SUBAPPLICATION logiBUS_AI_Calibrate_3P_OPC (* logiBUS_AI 3-Punkt-Kalibrierung, INI-persistiert, C_MIN/C_MID/C_MAX per Methode, alles per OPC-UA (ohne VT) *)
  (* Standard: 61499-2; Description: Copyright (c) 2026 Meisterschulen am Ostbahnhof This program and the accompanying materials are made available under the terms of the Eclipse Public License 2.0 which is available at https://www.eclipse.org/legal/epl-2.0/ SPDX-License-Identifier: EPL-2.0 *)
  (* Version 1.2, 2026-11-25, Franz Höpfinger, Meisterschulen am Ostbahnhof, SERVER_0 -> MyLib::net::SERVER_0_QO (IND nur bei QO=TRUE, RSP intern). Ein gescheitertes RSP meldet IND mit QO=FALSE, direkt IND->RSP ergab eine Endlosschleife. *)
  (* Version 1.1, 2026-11-04, Franz Höpfinger, Meisterschulen am Ostbahnhof, Neuer optionaler Ausgangs-Plug CAL_OUT (kalibrierter Wert = CALIBRATE.Y, AR) per AR_SPLIT_2 SplitCal zwischen CALIBRATE.Y und PublishCal - wie CAL_OUT in logiBUS_AI_Calibrate_3P_Remote_IDA_OPC. Damit kann z.B. ein Servo direkt am kalibrierten Wert haengen statt den eigenen OPC-UA-Knoten lokal zu abonnieren. Unverdrahtet lassen, wenn nicht gebraucht. *)
  (* Version 1.0, 2026-10-28, Franz Höpfinger, Meisterschulen am Ostbahnhof, Kopie von MyLib::sys::logiBUS_AI_Calibrate_3P_IDA_OPC (INIT-Kette Stand bf9ac7c9) ohne VT, fuer Stationen ohne VT (keine isobus_UT-Libs). InputRaw -> MyLib::sys::logiBUS_AI_Raw_AR_OPC, *_REF_LIT -> MyLib::sys::OPC_TO_AR2, Trigger* -> SERVER_0 (IND->RSP), Publish* -> MyLib::sys::AR_TO_Publish_OPC. VT-Objekt-Parameter entfallen, Kalibrierlogik und INI-Keys unveraendert. *)
  PACKAGE MyLib::sys;
  IMPORT logiBUS::io::AI::logiBUS_AI;
  IMPORT logiBUS::io::AI::logiBUS_AI_S;
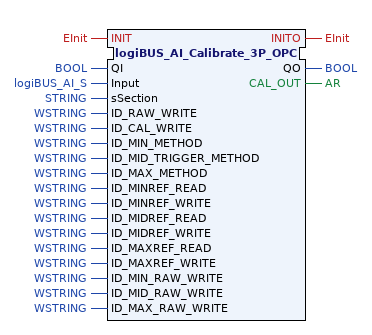
  EVENT_INPUT
    INIT : EInit; (* Initialization Request *)
  END_EVENT
  EVENT_OUTPUT
    INITO : EInit; (* Initialization Confirm *)
  END_EVENT
  VAR_INPUT
    QI : BOOL := TRUE; (* Quality Input - TRUE to enable service *)
    Input : logiBUS::io::AI::logiBUS_AI_S := logiBUS_AI::Invalid; (* Identify the Input AnalogInput_I1..I8 *)
    sSection : STRING; (* INI-Sektionsname fuer X_MIN/X_MID/X_MAX/MIN_REF/MID_REF/MAX_REF-Persistenz - pro Kanal eindeutig, sonst kollidieren die Kanaele in settings.ini *)
    ID_RAW_WRITE : WSTRING; (* Rohwert-Ruckmelde-Adresse (DWORD 0-4095, ACTION=PUBLISH) *)
    ID_CAL_WRITE : WSTRING; (* Kalibrierter-Wert-Ruckmelde-Adresse (REAL, ACTION=PUBLISH) *)
    ID_MIN_METHOD : WSTRING; (* Methodenadresse (ACTION=CREATE_METHOD) fuer den argumentlosen C_MIN-Trigger - gleichberechtigt zur lokalen VT-Taste aufrufbar, sowohl vom OPC-UA-Dashboard als auch per CLIENT_0 von einer anderen Station (siehe OPC_UA_VERNETZUNG.md Punkt 14 - kein Toggle/Subscribe-Umweg mehr) *)
    ID_MID_TRIGGER_METHOD : WSTRING; (* Methodenadresse (ACTION=CREATE_METHOD) fuer den argumentlosen C_MID-Trigger - siehe ID_MIN_METHOD *)
    ID_MAX_METHOD : WSTRING; (* Methodenadresse (ACTION=CREATE_METHOD) fuer den argumentlosen C_MAX-Trigger - siehe ID_MIN_METHOD *)
    ID_MINREF_READ : WSTRING; (* Remote-Subscribe-Adresse MIN_REF-Referenzwert (REAL, ACTION=SUBSCRIBE) *)
    ID_MINREF_WRITE : WSTRING; (* Remote-Echo-Adresse MIN_REF-Referenzwert (REAL, ACTION=PUBLISH) *)
    ID_MIDREF_READ : WSTRING; (* Remote-Subscribe-Adresse MID_REF-Referenzwert (REAL, ACTION=SUBSCRIBE) *)
    ID_MIDREF_WRITE : WSTRING; (* Remote-Echo-Adresse MID_REF-Referenzwert (REAL, ACTION=PUBLISH) *)
    ID_MAXREF_READ : WSTRING; (* Remote-Subscribe-Adresse MAX_REF-Referenzwert (REAL, ACTION=SUBSCRIBE) *)
    ID_MAXREF_WRITE : WSTRING; (* Remote-Echo-Adresse MAX_REF-Referenzwert (REAL, ACTION=PUBLISH) *)
    ID_MIN_RAW_WRITE : WSTRING; (* Rohwert-am-MIN-Kalibrierpunkt-Publish-Adresse (REAL, ACTION=PUBLISH) *)
    ID_MID_RAW_WRITE : WSTRING; (* Rohwert-am-MID-Kalibrierpunkt-Publish-Adresse (REAL, ACTION=PUBLISH) *)
    ID_MAX_RAW_WRITE : WSTRING; (* Rohwert-am-MAX-Kalibrierpunkt-Publish-Adresse (REAL, ACTION=PUBLISH) *)
  END_VAR
  VAR_OUTPUT
    QO : BOOL; (* Quality Output - TRUE if service executed successfully *)
  END_VAR
  PLUGS
    CAL_OUT : adapter::types::unidirectional::AR; (* Optional: kalibrierter Wert (= CALIBRATE.Y) fuer externe Consumer, statt eigenem lokalen OPC-UA-Self-Subscribe auf ID_CAL_WRITE. Unverdrahtet lassen, wenn nicht gebraucht. *)
  END_PLUGS
  FBS
    CALIBRATE : adapter::Engineering::measurements::AR_CALIBRATE_3P_REF(xClipping := FALSE);
    INI_X_MIN : eclipse4diac::storage::INI_AR2(SETM := TRUE, KEY := 'X_MIN', DEFAULT_VALUE := REAL#0.0);
    INI_X_MID : eclipse4diac::storage::INI_AR2(SETM := TRUE, KEY := 'X_MID', DEFAULT_VALUE := REAL#0.0);
    INI_X_MAX : eclipse4diac::storage::INI_AR2(SETM := TRUE, KEY := 'X_MAX', DEFAULT_VALUE := REAL#0.0);
    INI_MIN_REF : eclipse4diac::storage::INI_AR2(SETM := TRUE, KEY := 'MIN_REF', DEFAULT_VALUE := REAL#-100.0);
    INI_MID_REF : eclipse4diac::storage::INI_AR2(SETM := TRUE, KEY := 'MID_REF', DEFAULT_VALUE := REAL#0.0);
    INI_MAX_REF : eclipse4diac::storage::INI_AR2(SETM := TRUE, KEY := 'MAX_REF', DEFAULT_VALUE := REAL#100.0);
    TapMinRaw : adapter::events::bidirectional::AR2_SPLIT_FWD_REV;
    TapMidRaw : adapter::events::bidirectional::AR2_SPLIT_FWD_REV;
    TapMaxRaw : adapter::events::bidirectional::AR2_SPLIT_FWD_REV;
    AND_QO : iec61131::booleanOperators::AND_BOOL_18;
    SplitCal : adapter::events::unidirectional::AR_SPLIT_2;
  END_FBS
  SUBAPPS
    InputRaw : MyLib::sys::logiBUS_AI_Raw_AR_OPC;
    MIN_REF_LIT : MyLib::sys::OPC_TO_AR2;
    MID_REF_LIT : MyLib::sys::OPC_TO_AR2;
    MAX_REF_LIT : MyLib::sys::OPC_TO_AR2;
    TriggerMIN : MyLib::net::SERVER_0_QO; (* RSP direkt auf IND (sonst 4s Server-Lock) *)
    TriggerMID : MyLib::net::SERVER_0_QO; (* RSP direkt auf IND (sonst 4s Server-Lock) *)
    TriggerMAX : MyLib::net::SERVER_0_QO; (* RSP direkt auf IND (sonst 4s Server-Lock) *)
    PublishCal : MyLib::sys::AR_TO_Publish_OPC;
    PublishMinRaw : MyLib::sys::AR_TO_Publish_OPC;
    PublishMidRaw : MyLib::sys::AR_TO_Publish_OPC;
    PublishMaxRaw : MyLib::sys::AR_TO_Publish_OPC;
  END_SUBAPPS
  EVENT_CONNECTIONS
    TriggerMIN.IND TO CALIBRATE.C_MIN;
    TriggerMID.IND TO CALIBRATE.C_MID;
    TriggerMAX.IND TO CALIBRATE.C_MAX;
    INIT TO TriggerMIN.INIT;
    CALIBRATE.INITO TO PublishCal.INIT;
    INI_X_MIN.INITO TO INI_X_MID.INIT;
    INI_X_MID.INITO TO INI_X_MAX.INIT;
    INI_X_MAX.INITO TO INI_MIN_REF.INIT;
    INI_MIN_REF.INITO TO INI_MID_REF.INIT;
    INI_MID_REF.INITO TO INI_MAX_REF.INIT;
    InputRaw.INITO TO MIN_REF_LIT.INIT;
    MIN_REF_LIT.INITO TO MID_REF_LIT.INIT;
    MID_REF_LIT.INITO TO MAX_REF_LIT.INIT;
    TriggerMIN.INITO TO TriggerMID.INIT;
    TriggerMID.INITO TO TriggerMAX.INIT;
    PublishCal.INITO TO PublishMinRaw.INIT;
    PublishMinRaw.INITO TO PublishMidRaw.INIT;
    PublishMidRaw.INITO TO PublishMaxRaw.INIT;
    INI_MAX_REF.INITO TO INITO;
    INI_MAX_REF.INITO TO AND_QO.REQ;
    TriggerMAX.INITO TO InputRaw.INIT;
    MAX_REF_LIT.INITO TO CALIBRATE.INIT;
    PublishMaxRaw.INITO TO INI_X_MIN.INIT;
  END_CONNECTIONS
  DATA_CONNECTIONS
    Input TO InputRaw.Input;
    sSection TO INI_X_MIN.SECTION;
    sSection TO INI_X_MID.SECTION;
    sSection TO INI_X_MAX.SECTION;
    sSection TO INI_MIN_REF.SECTION;
    sSection TO INI_MID_REF.SECTION;
    sSection TO INI_MAX_REF.SECTION;
    ID_RAW_WRITE TO InputRaw.ID_RAW_WRITE;
    ID_CAL_WRITE TO PublishCal.ID_WRITE;
    ID_MIN_METHOD TO TriggerMIN.ID;
    ID_MID_TRIGGER_METHOD TO TriggerMID.ID;
    ID_MAX_METHOD TO TriggerMAX.ID;
    ID_MINREF_READ TO MIN_REF_LIT.ID_READ;
    ID_MINREF_WRITE TO MIN_REF_LIT.ID_WRITE;
    ID_MIDREF_READ TO MID_REF_LIT.ID_READ;
    ID_MIDREF_WRITE TO MID_REF_LIT.ID_WRITE;
    ID_MAXREF_READ TO MAX_REF_LIT.ID_READ;
    ID_MAXREF_WRITE TO MAX_REF_LIT.ID_WRITE;
    ID_MIN_RAW_WRITE TO PublishMinRaw.ID_WRITE;
    ID_MID_RAW_WRITE TO PublishMidRaw.ID_WRITE;
    ID_MAX_RAW_WRITE TO PublishMaxRaw.ID_WRITE;
    QI TO CALIBRATE.QI;
    QI TO INI_X_MIN.QI;
    QI TO INI_X_MID.QI;
    QI TO INI_X_MAX.QI;
    QI TO INI_MIN_REF.QI;
    QI TO INI_MID_REF.QI;
    QI TO INI_MAX_REF.QI;
    QI TO InputRaw.QI;
    QI TO MIN_REF_LIT.QI;
    QI TO MID_REF_LIT.QI;
    QI TO MAX_REF_LIT.QI;
    QI TO TriggerMIN.QI;
    QI TO TriggerMID.QI;
    QI TO TriggerMAX.QI;
    QI TO PublishCal.QI;
    QI TO PublishMinRaw.QI;
    QI TO PublishMidRaw.QI;
    QI TO PublishMaxRaw.QI;
    CALIBRATE.QO TO AND_QO.IN1;
    INI_X_MIN.QO TO AND_QO.IN2;
    INI_X_MID.QO TO AND_QO.IN3;
    INI_X_MAX.QO TO AND_QO.IN4;
    INI_MIN_REF.QO TO AND_QO.IN5;
    INI_MID_REF.QO TO AND_QO.IN6;
    INI_MAX_REF.QO TO AND_QO.IN7;
    InputRaw.QO TO AND_QO.IN8;
    MIN_REF_LIT.QO TO AND_QO.IN9;
    MID_REF_LIT.QO TO AND_QO.IN10;
    MAX_REF_LIT.QO TO AND_QO.IN11;
    TriggerMIN.QO TO AND_QO.IN12;
    TriggerMID.QO TO AND_QO.IN13;
    TriggerMAX.QO TO AND_QO.IN14;
    PublishCal.QO TO AND_QO.IN15;
    PublishMinRaw.QO TO AND_QO.IN16;
    PublishMidRaw.QO TO AND_QO.IN17;
    PublishMaxRaw.QO TO AND_QO.IN18;
    AND_QO.OUT TO QO;
  END_CONNECTIONS
  ADAPTER_CONNECTIONS
    InputRaw.AR_OUT TO CALIBRATE.X;
    CALIBRATE.X_MIN TO TapMinRaw.IN;
    TapMinRaw.OUT TO INI_X_MIN.VAL;
    TapMinRaw.REV_OUT TO PublishMinRaw.AR_IN;
    CALIBRATE.X_MID TO TapMidRaw.IN;
    TapMidRaw.OUT TO INI_X_MID.VAL;
    TapMidRaw.REV_OUT TO PublishMidRaw.AR_IN;
    CALIBRATE.X_MAX TO TapMaxRaw.IN;
    TapMaxRaw.OUT TO INI_X_MAX.VAL;
    TapMaxRaw.REV_OUT TO PublishMaxRaw.AR_IN;
    CALIBRATE.MIN_REF TO INI_MIN_REF.VAL;
    CALIBRATE.MID_REF TO INI_MID_REF.VAL;
    CALIBRATE.MAX_REF TO INI_MAX_REF.VAL;
    MIN_REF_LIT.VALUEO TO CALIBRATE.Y_MIN;
    MID_REF_LIT.VALUEO TO CALIBRATE.Y_MID;
    MAX_REF_LIT.VALUEO TO CALIBRATE.Y_MAX;
    CALIBRATE.Y TO SplitCal.IN;
    SplitCal.OUT1 TO PublishCal.AR_IN;
    SplitCal.OUT2 TO CAL_OUT;
  END_CONNECTIONS
END_SUBAPPLICATION
